(* Logix 5000 project; controller TFF vendor 1 type 14 code 107 rev 34.11; software revision 34.03; part 27 of 36 *)
(* tags used below, declared in another part *)
   BufferSteps0_Prev : STRING25;
   Config : Configuration;   // Index Array used in configuration routines
   Index : DINT;   // Index
   RecipeStepLog_DateTime_Empty : STRING25;   // Empty String
   RecipeStepLog_DateTime_Log : STRING25;   // Last Date Time received from HMI
   RecipeStepLog_DateTime_Prev : STRING25;
   RecipeStepLog_Timer : TIMER;   // RecipeStepLog Watchdog Timer
   AI101 : ALIAS FOR AnalogPoint[10];   // Filtrate Conductivity
   AI101_SIG : ALIAS FOR DigitalPoint[90];
   AI102 : ALIAS FOR AnalogPoint[11];   // Filtrate UV
   AI102_SIG : ALIAS FOR DigitalPoint[91];
   AI103 : ALIAS FOR AnalogPoint[12];   // Filtrate UV
   AI103_SIG : ALIAS FOR DigitalPoint[92];
   AI104 : ALIAS FOR AnalogPoint[9];   // Filtrate pH
   AI104_SIG : ALIAS FOR DigitalPoint[105];
   CCPSystem : CCPSystem;   // CCP System Data
   DigitalInput : BOOL[256];   // Digital Input Array these bits are copied from Input cards.
   DigitalPoint : DigitalPoint[150];   // Digital Point Array
   ES001 : ALIAS FOR DigitalPoint[3];   // Emergency Stop
   FI003 : ALIAS FOR AnalogPoint[17];
   FI003_SIG : ALIAS FOR DigitalPoint[106];
   FI101 : ALIAS FOR AnalogPoint[2];   // Filtrate Flow
   FI101_SIG : ALIAS FOR DigitalPoint[93];
   HTCCollectorError : BOOL;   // Hist. Data Collect. Error
   HTCHeartBeat : BOOL;   // Historical Data Collection heartbeat (Set to 1 by HMI Reset to 0 by PLC)
   MIX001 : ALIAS FOR AnalogPoint[14];   // Mixer Speed
   MIX001_SIG : ALIAS FOR DigitalPoint[104];
   Mixer : Mixer;   // Mixer config. structure
   OperatingTime : OperatingTime;
   Options : Options;   // Options List
   PcToPLCHeartBeat : BOOL;   // PC to PLC communication heartbeat Set to 1 by HMI Reset to 0 by plc
   PCV001 : ALIAS FOR AnalogPoint[3];   // Retentate Pressure Control Valve Position
   PCV001_SIG : ALIAS FOR DigitalPoint[102];
   PCV101 : ALIAS FOR AnalogPoint[4];   // Filtrate Pressure Control Valve Position
   PCV101_SIG : ALIAS FOR DigitalPoint[103];
   Phase0 : ALIAS FOR Phase[0];   // Phase 0
   PI001 : ALIAS FOR AnalogPoint[5];   // Feed Pressure
   PI001_SIG : ALIAS FOR DigitalPoint[97];
   PI002 : ALIAS FOR AnalogPoint[6];   // Retentate Pressure
   PI002_SIG : ALIAS FOR DigitalPoint[98];
   PI101 : ALIAS FOR AnalogPoint[7];   // Filtrate Pressure
   PI101_SIG : ALIAS FOR DigitalPoint[99];
   PI401 : ALIAS FOR AnalogPoint[8];   // Transfer Pump Pressure
   PI401_SIG : ALIAS FOR DigitalPoint[100];
   PSH001 : ALIAS FOR DigitalPoint[4];   // Feed Pump High Pressure
   PSH401 : ALIAS FOR DigitalPoint[5];   // Transfer Pump High Pressure
   PSL603 : ALIAS FOR DigitalPoint[10];   // Manifold Valves Air Defect
   Rack_Murr_Node0_Smart : IO_Station;   // Status of Node 0 Smart
   Rack_Murr_Node1_TF2S : IO_Station;   // Status of Node 1 TF2S
   Rack_Murr_Node1_TF3S : IO_Station;   // Status of Node 1 TF3S
   Rack_Murr_Node3_PUMP : IO_Station;   // Status of Node 3 Pump
   Rack_Murr_Node4_Instrum_TFF1 : IO_Station;   // Status of Node 4 Instrum TFF1
   Rack_Murr_Node4_Instrum_TFF2 : IO_Station;   // Status of Node 4 Instrum TFF2
   Rack_Murr_Node4_Instrum_TFF3 : IO_Station;   // Status of Node 4 Instrum TFF3
   Rack_Murr_Node4_Instrum_TFF4 : IO_Station;   // Status of Node 4 Instrum TFF4
   Rack_Murr_Node4_Instrum_TFF5 : IO_Station;   // Status of Node 4 Instrum TFF5
   Rack_Murr_Node5_Tank100 : IO_Station;   // Status of Node 5 Tank 100L
   Rack_Murr_Node5_Tank250 : IO_Station;   // Status of Node 5 Tank 250L
   Rack_Murr_Node5_Tank50 : IO_Station;   // Status of Node 5 Tank 50L
   Rack_Murr_Node6_IND331_WI001 : IO_Station;   // Status of Node 6 IND331 WI001
   Rack_Murr_Node7_IND131_WI101 : IO_Station;   // Status of Node 7 IND131 WI101
   RecipeStepLog_DateTime : STRING25;
   SIC001DF : ALIAS FOR DigitalPoint[8];   // Feed Pump Defect
   SIC002DF : ALIAS FOR DigitalPoint[9];   // Transfer Pump Defect
   SIC003DF : ALIAS FOR DigitalPoint[14];   // Mixer Defect
   SRL001 : ALIAS FOR DigitalPoint[15];   // Tank Skid Remote / Standalone
   Tank : TankManagement;   // Tank Management
   ThisSystem : SystemType;
   TI001 : ALIAS FOR AnalogPoint[13];   // Feed Bag Temperature
   TI001_SIG : ALIAS FOR DigitalPoint[101];
   WI001 : ALIAS FOR AnalogPoint[15];   // Feed Bag Weight
   WI001_SIG : ALIAS FOR DigitalPoint[94];
   WI101 : ALIAS FOR AnalogPoint[0];   // Filtrate Weight
   WI101_SIG : ALIAS FOR DigitalPoint[95];
   WI102 : ALIAS FOR AnalogPoint[1];   // Customer Filtrate Weight
   WI102_SIG : ALIAS FOR DigitalPoint[96];
   XC102_3DF : ALIAS FOR DigitalPoint[13];   // C8000 Defect
   XS001 : ALIAS FOR DigitalPoint[1];   // Door Closed
   XS002 : ALIAS FOR DigitalPoint[6];   // Clamshell Locking 1 Closed
   XS003 : ALIAS FOR DigitalPoint[7];   // Clamshell Locking 2 Closed
   XS006 : ALIAS FOR DigitalPoint[2];   // Door to Frame Locking Closed
   XS011 : ALIAS FOR DigitalPoint[11];   // Pump P001 Type
   XS012 : ALIAS FOR DigitalPoint[12];   // Pump P002 Type
   YA01 : ALIAS FOR DigitalPoint[50];   // PC to PLC communication failure
   YA02 : ALIAS FOR DigitalPoint[51];   // CCP Runtime communication failure
   YA03 : ALIAS FOR DigitalPoint[52];   // Historical Data collection failure
   YA06 : ALIAS FOR DigitalPoint[55];   // Node 0 communication failure - Smart
   YA07 : ALIAS FOR DigitalPoint[56];   // Node 0 internal defect - Smart
   YA08 : ALIAS FOR DigitalPoint[57];   // Node 1 communication failure - Clamshell
   YA09 : ALIAS FOR DigitalPoint[58];   // Node 1 internal defect - Clamshell
   YA13 : ALIAS FOR DigitalPoint[62];   // Tank Size Mismatch
   YA14 : ALIAS FOR DigitalPoint[63];   // SQL Server Write Failure
   YA15 : ALIAS FOR DigitalPoint[69];   // Node 3 Communication Failure - Pump
   YA16 : ALIAS FOR DigitalPoint[70];   // Node 3 Internal Defect - Pump
   YA17 : ALIAS FOR DigitalPoint[71];   // Node 4 Communication Failure - Instrum
   YA18 : ALIAS FOR DigitalPoint[72];   // Node 4 Internal Defect - Instrum
   YA19 : ALIAS FOR DigitalPoint[73];   // Node 5 Communication Failure - Tank
   YA20 : ALIAS FOR DigitalPoint[74];   // Node 5 Internal Defect - Tank
   YA21 : ALIAS FOR DigitalPoint[75];   // Node 6 IND331 Communication Failure
   YA22 : ALIAS FOR DigitalPoint[76];   // Node 7 IND131 Communication Failure
   YA41 : ALIAS FOR DigitalPoint[77];   // YA41 Operating Time Exceeded
   ZSDF : ALIAS FOR DigitalPoint[68];   // ZSDF Clamshell Locking Defect
(* Process, continued *)

ROUTINE InputDigitalPoint   (* ladder *)
// Digital Point Routine
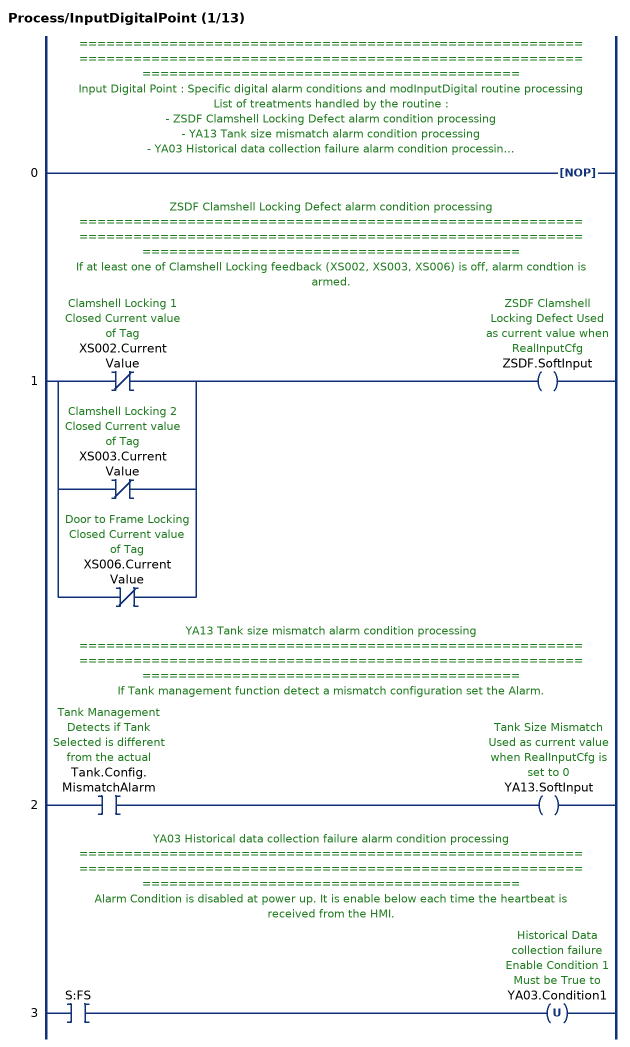
   // ==========================================================================================================================================================
   //                                                                                   Input Digital Point : Specific digital alarm conditions and modInputDigital routine processing
   //                                                     List of treatments handled by the routine :
   //                                                          - ZSDF Clamshell Locking Defect alarm condition processing
   //                                                          - YA13 Tank size mismatch alarm condition processing
   //                                                          - YA03 Historical data collection failure alarm condition processing
   //                                                          - YA01 PC to PLC com. failure alarm condition processing
   //                                                          - YA02 CCP Runtime com. failure alarm condition processing
   //                                                          - YA14 SQL Write failure alarm condition processing
   //                                                          - Node 0 communication failure and internal defect (YA06 and YA07)
   //                                                          - Node 1 communication failure and internal defect (YA08 and YA09)
   //                                                          - Node 3 communication failure and internal defect (YA15 and YA16)
   //                                                          - Node 4 communication failure and internal defect (YA17 and YA18)
   //                                                          - Node 5 communication failure and internal defect (YA19 and YA20)
   //                                                          - IND331 communication failure and internal defect (YA21)
   //                                                          - IND131 communication failure and internal defect (YA22)
   //                               - YA41 Operating Time Exceeded (YA41)
   //                                                          - Analog Signal Failure
   //                                                          - modInputDigital Loop
   //                                                     -----------------------------------------------------------------------------------------------------------------------------------------------------
   //                                                     History
   //                                            2019-AUG-13 - Actemium - B. Roch - Initial version for Candidate Release 3.00.00.00.a
   //                              2019-SEP-25 - Actemium - B. Roch - Modification for Candidate Release 3.00.00.00
   // - Add condition to comput SQL Write failure alarm (not in step 1)
   //                                 2020-SEP-14 - Merck - Q. Spindler - Modifications for Candidate Release 3.00.00.01.a
   //                                                   - Add Conditions to YA20, YA18, and YA09 so only connected nodes can trigger internal deffect
   //  - Change YA14 Alarm condition processing to add HMI Watchdog
   // - Add FI003_SIG
   // 2021-MAY-28 - DAVIDSON- Ch. ARBOGAST - Modifications for Candidate Release 3.01.00.00.a
   //  - Rung 6 unlatch YA03: add test not HTCColletorError (new tag - bool)
   //  - Add rung 30: write YA41.softInput - DigitalPoint[77] - Operating Time Exceeded
   // 2023-MAR-29 - DAVIDSON- Ch. ARBOGAST - Modifications for Candidate Release 3.02.00.00.a
   //  - Rung 2; replace DigitalPoint[41].SoftInput by YA13.SoftInput
   // ==========================================================================================================================================================
   0: NOP();
   // ZSDF Clamshell Locking Defect alarm condition processing
   // ==========================================================================================================================================================
   // If at least one of Clamshell Locking feedback (XS002, XS003, XS006) is off, alarm condtion is armed.
   1: [XIO(XS002.CurrentValue) ,XIO(XS003.CurrentValue) ,XIO(XS006.CurrentValue) ]OTE(ZSDF.SoftInput);
   // YA13 Tank size mismatch alarm condition processing
   // ==========================================================================================================================================================
   // If Tank management function detect a mismatch configuration set the Alarm.
   2: XIC(Tank.Config.MismatchAlarm)OTE(YA13.SoftInput);
   // YA03 Historical data collection failure alarm condition processing
   // ==========================================================================================================================================================
   // Alarm Condition is disabled at power up. It is enable below each time the heartbeat is received from the HMI.
   3: XIC(S:FS)OTU(YA03.Condition1);
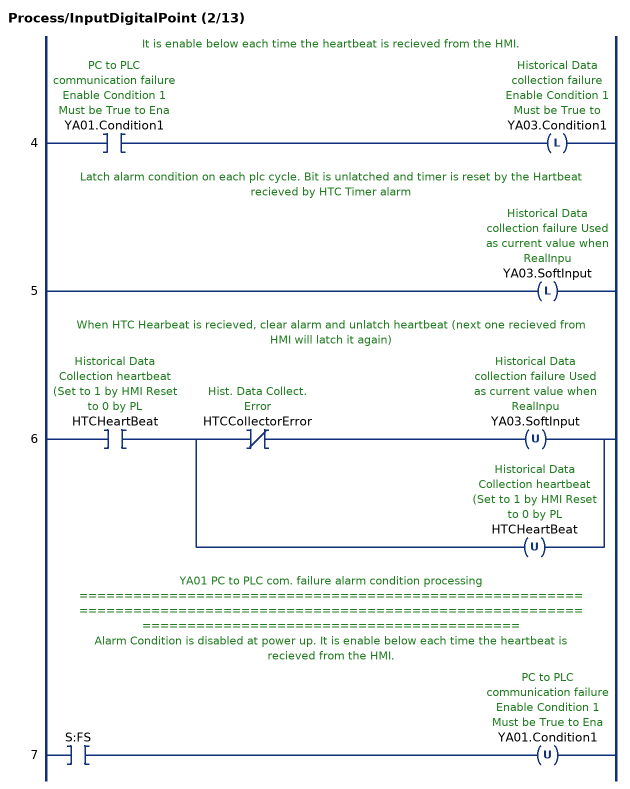
   // It is enable below each time the heartbeat is recieved from the HMI.
   4: XIC(YA01.Condition1)OTL(YA03.Condition1);
   // Latch alarm condition on each plc cycle. Bit is unlatched and timer is reset by the Hartbeat recieved by HTC Timer alarm
   5: OTL(YA03.SoftInput);
   // When HTC Hearbeat is recieved, clear alarm and unlatch heartbeat (next one recieved from HMI will latch it again)
   6: XIC(HTCHeartBeat)[XIO(HTCCollectorError) OTU(YA03.SoftInput) ,OTU(HTCHeartBeat) ];
   // YA01 PC to PLC com. failure alarm condition processing
   // ==========================================================================================================================================================
   // Alarm Condition is disabled at power up. It is enable below each time the heartbeat is recieved from the HMI.
   7: XIC(S:FS)OTU(YA01.Condition1);
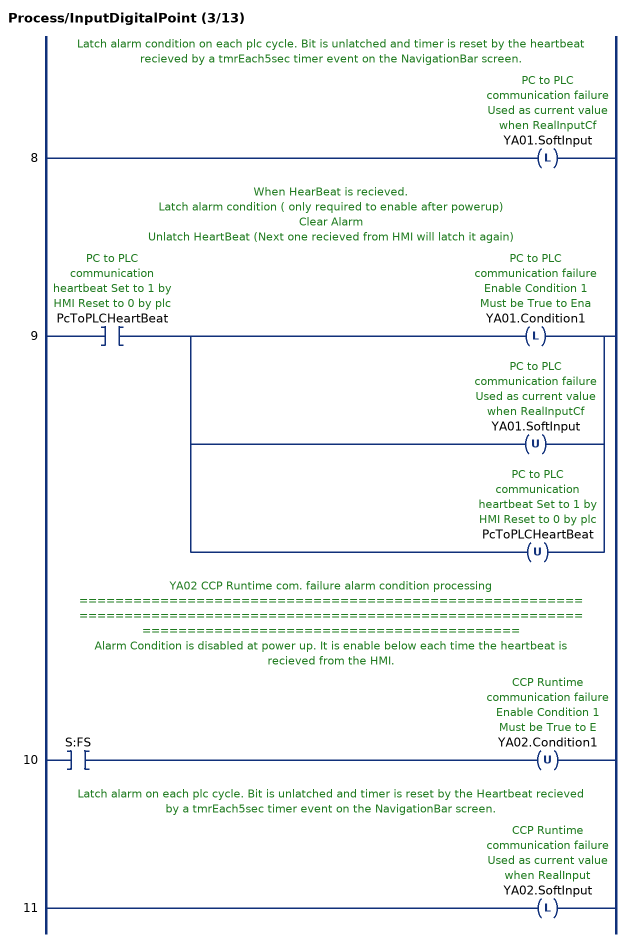
   // Latch alarm condition on each plc cycle. Bit is unlatched and timer is reset by the heartbeat recieved by a tmrEach5sec timer event on the NavigationBar screen.
   8: OTL(YA01.SoftInput);
   // When HearBeat is recieved.
   //         Latch alarm condition ( only required to enable after powerup)
   //         Clear Alarm
   //        Unlatch HeartBeat (Next one recieved from HMI will latch it again)
   9: XIC(PcToPLCHeartBeat)[OTL(YA01.Condition1) ,OTU(YA01.SoftInput) ,OTU(PcToPLCHeartBeat) ];
   // YA02 CCP Runtime com. failure alarm condition processing
   // ==========================================================================================================================================================
   // Alarm Condition is disabled at power up. It is enable below each time the heartbeat is recieved from the HMI.
   10: XIC(S:FS)OTU(YA02.Condition1);
   // Latch alarm on each plc cycle. Bit is unlatched and timer is reset by the Heartbeat recieved by a tmrEach5sec timer event on the NavigationBar screen.
   11: OTL(YA02.SoftInput);
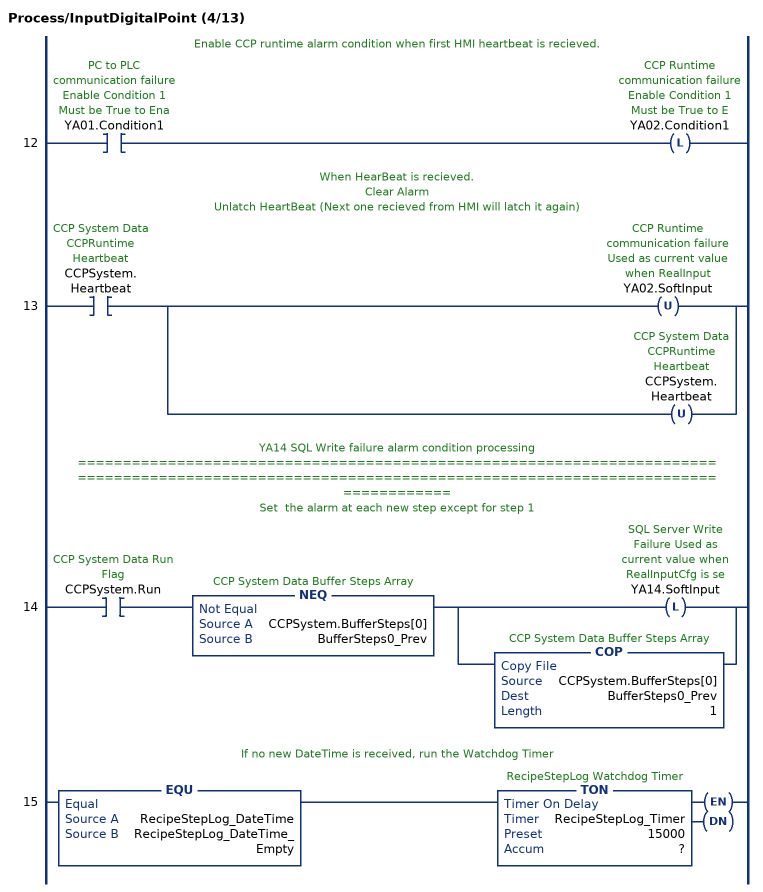
   // Enable CCP runtime alarm condition when first HMI heartbeat is recieved.
   12: XIC(YA01.Condition1)OTL(YA02.Condition1);
   // When HearBeat is recieved.
   //         Clear Alarm
   //        Unlatch HeartBeat (Next one recieved from HMI will latch it again)
   13: XIC(CCPSystem.Heartbeat)[OTU(YA02.SoftInput) ,OTU(CCPSystem.Heartbeat) ];
   // YA14 SQL Write failure alarm condition processing
   // ==========================================================================================================================================================
   // Set  the alarm at each new step except for step 1
   14: XIC(CCPSystem.Run)NEQ(CCPSystem.BufferSteps[0],BufferSteps0_Prev)[OTL(YA14.SoftInput) ,COP(CCPSystem.BufferSteps[0],BufferSteps0_Prev,1) ];
   // If no new DateTime is received, run the Watchdog Timer
   15: EQU(RecipeStepLog_DateTime,RecipeStepLog_DateTime_Empty)TON(RecipeStepLog_Timer,?,?);
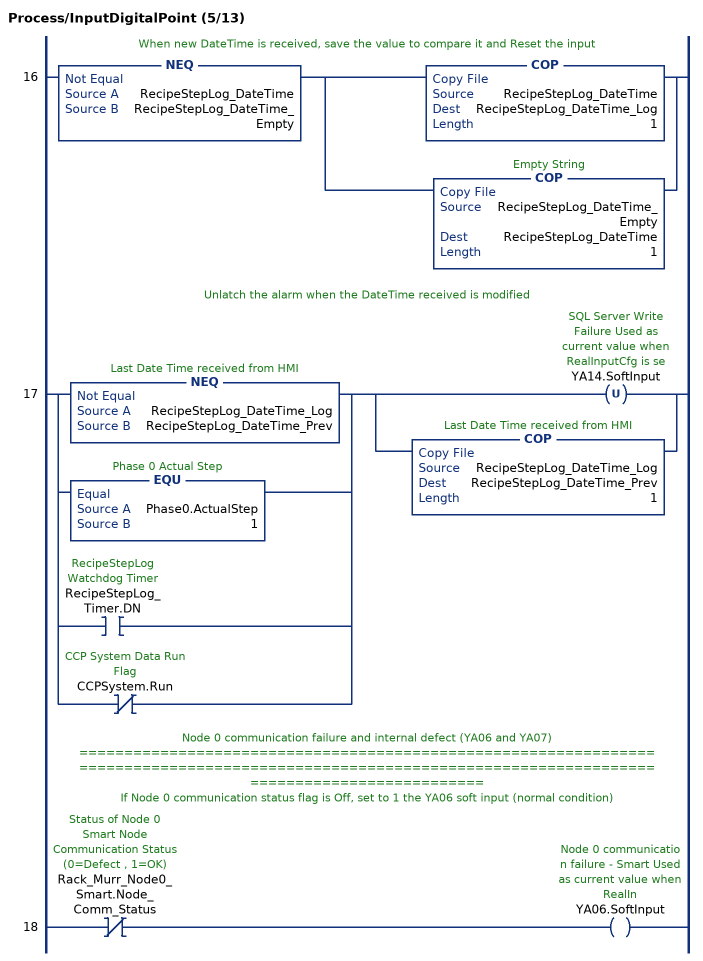
   // When new DateTime is received, save the value to compare it and Reset the input
   16: NEQ(RecipeStepLog_DateTime,RecipeStepLog_DateTime_Empty)[COP(RecipeStepLog_DateTime,RecipeStepLog_DateTime_Log,1) ,COP(RecipeStepLog_DateTime_Empty,RecipeStepLog_DateTime,1) ];
   // Unlatch the alarm when the DateTime received is modified
   17: [NEQ(RecipeStepLog_DateTime_Log,RecipeStepLog_DateTime_Prev) ,EQU(Phase0.ActualStep,1) ,XIC(RecipeStepLog_Timer.DN) ,XIO(CCPSystem.Run) ][OTU(YA14.SoftInput) ,COP(RecipeStepLog_DateTime_Log,RecipeStepLog_DateTime_Prev,1) ];
   // Node 0 communication failure and internal defect (YA06 and YA07)
   // ==========================================================================================================================================================
   // If Node 0 communication status flag is Off, set to 1 the YA06 soft input (normal condition)
   18: XIO(Rack_Murr_Node0_Smart.Node_Comm_Status)OTE(YA06.SoftInput);
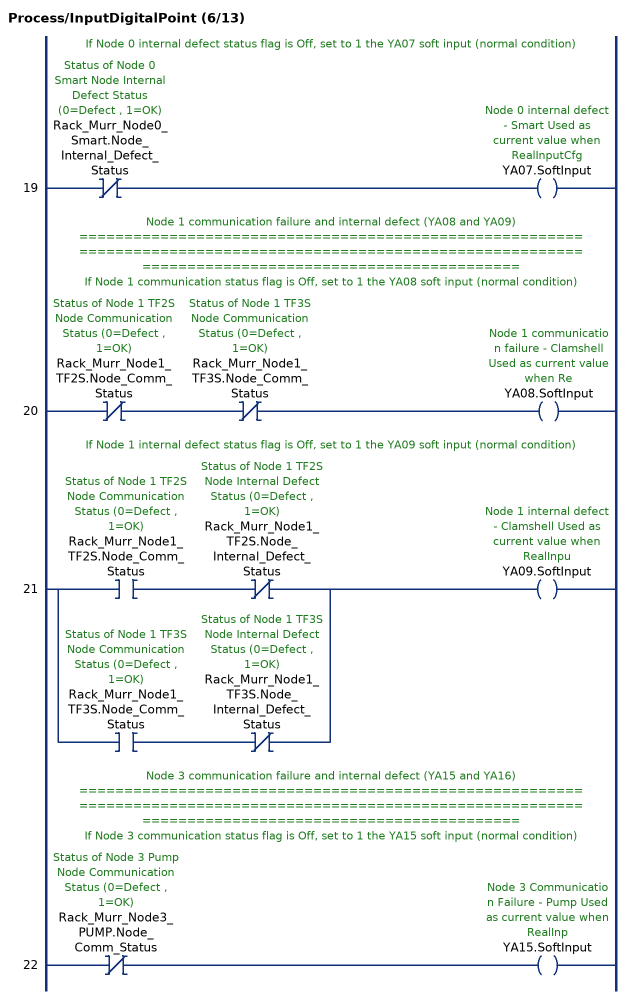
   // If Node 0 internal defect status flag is Off, set to 1 the YA07 soft input (normal condition)
   19: XIO(Rack_Murr_Node0_Smart.Node_Internal_Defect_Status)OTE(YA07.SoftInput);
   // Node 1 communication failure and internal defect (YA08 and YA09)
   // ==========================================================================================================================================================
   // If Node 1 communication status flag is Off, set to 1 the YA08 soft input (normal condition)
   20: XIO(Rack_Murr_Node1_TF2S.Node_Comm_Status)XIO(Rack_Murr_Node1_TF3S.Node_Comm_Status)OTE(YA08.SoftInput);
   // If Node 1 internal defect status flag is Off, set to 1 the YA09 soft input (normal condition)
   21: [XIC(Rack_Murr_Node1_TF2S.Node_Comm_Status) XIO(Rack_Murr_Node1_TF2S.Node_Internal_Defect_Status) ,XIC(Rack_Murr_Node1_TF3S.Node_Comm_Status) XIO(Rack_Murr_Node1_TF3S.Node_Internal_Defect_Status) ]OTE(YA09.SoftInput);
   // Node 3 communication failure and internal defect (YA15 and YA16)
   // ==========================================================================================================================================================
   // If Node 3 communication status flag is Off, set to 1 the YA15 soft input (normal condition)
   22: XIO(Rack_Murr_Node3_PUMP.Node_Comm_Status)OTE(YA15.SoftInput);
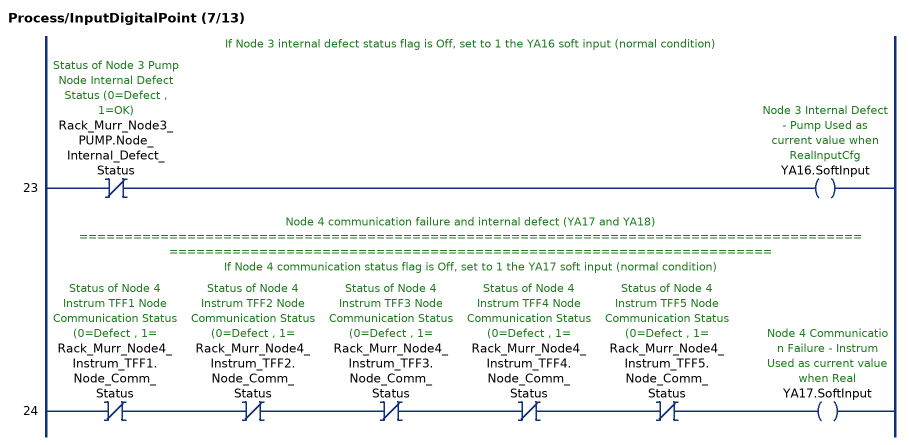
   // If Node 3 internal defect status flag is Off, set to 1 the YA16 soft input (normal condition)
   23: XIO(Rack_Murr_Node3_PUMP.Node_Internal_Defect_Status)OTE(YA16.SoftInput);
   // Node 4 communication failure and internal defect (YA17 and YA18)
   // ==========================================================================================================================================================
   // If Node 4 communication status flag is Off, set to 1 the YA17 soft input (normal condition)
   24: XIO(Rack_Murr_Node4_Instrum_TFF1.Node_Comm_Status)XIO(Rack_Murr_Node4_Instrum_TFF2.Node_Comm_Status)XIO(Rack_Murr_Node4_Instrum_TFF3.Node_Comm_Status)XIO(Rack_Murr_Node4_Instrum_TFF4.Node_Comm_Status)XIO(Rack_Murr_Node4_Instrum_TFF5.Node_Comm_Status)OTE(YA17.SoftInput);
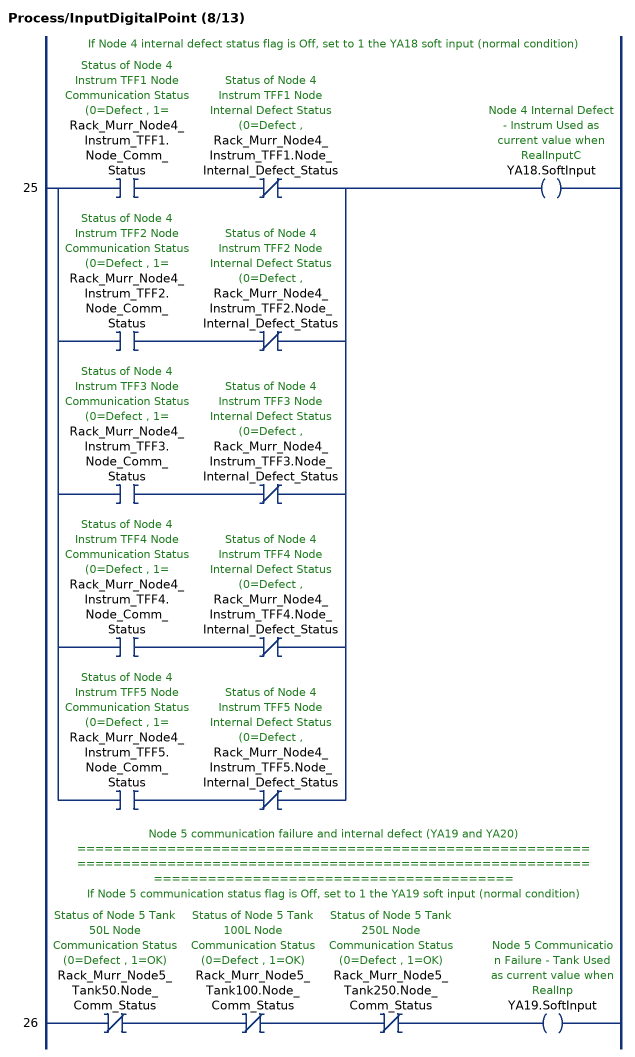
   // If Node 4 internal defect status flag is Off, set to 1 the YA18 soft input (normal condition)
   25: [XIC(Rack_Murr_Node4_Instrum_TFF1.Node_Comm_Status) XIO(Rack_Murr_Node4_Instrum_TFF1.Node_Internal_Defect_Status) ,XIC(Rack_Murr_Node4_Instrum_TFF2.Node_Comm_Status) XIO(Rack_Murr_Node4_Instrum_TFF2.Node_Internal_Defect_Status) ,XIC(Rack_Murr_Node4_Instrum_TFF3.Node_Comm_Status) XIO(Rack_Murr_Node4_Instrum_TFF3.Node_Internal_Defect_Status) ,XIC(Rack_Murr_Node4_Instrum_TFF4.Node_Comm_Status) XIO(Rack_Murr_Node4_Instrum_TFF4.Node_Internal_Defect_Status) ,XIC(Rack_Murr_Node4_Instrum_TFF5.Node_Comm_Status) XIO(Rack_Murr_Node4_Instrum_TFF5.Node_Internal_Defect_Status) ]OTE(YA18.SoftInput);
   // Node 5 communication failure and internal defect (YA19 and YA20)
   // ==========================================================================================================================================================
   // If Node 5 communication status flag is Off, set to 1 the YA19 soft input (normal condition)
   26: XIO(Rack_Murr_Node5_Tank50.Node_Comm_Status)XIO(Rack_Murr_Node5_Tank100.Node_Comm_Status)XIO(Rack_Murr_Node5_Tank250.Node_Comm_Status)OTE(YA19.SoftInput);
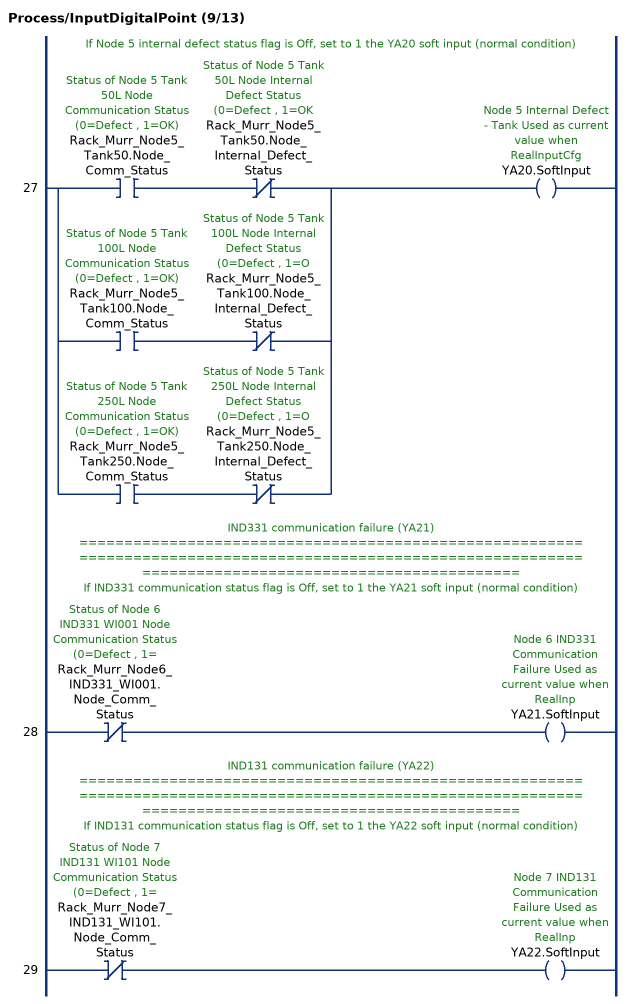
   // If Node 5 internal defect status flag is Off, set to 1 the YA20 soft input (normal condition)
   27: [XIC(Rack_Murr_Node5_Tank50.Node_Comm_Status) XIO(Rack_Murr_Node5_Tank50.Node_Internal_Defect_Status) ,XIC(Rack_Murr_Node5_Tank100.Node_Comm_Status) XIO(Rack_Murr_Node5_Tank100.Node_Internal_Defect_Status) ,XIC(Rack_Murr_Node5_Tank250.Node_Comm_Status) XIO(Rack_Murr_Node5_Tank250.Node_Internal_Defect_Status) ]OTE(YA20.SoftInput);
   // IND331 communication failure (YA21)
   // ==========================================================================================================================================================
   // If IND331 communication status flag is Off, set to 1 the YA21 soft input (normal condition)
   28: XIO(Rack_Murr_Node6_IND331_WI001.Node_Comm_Status)OTE(YA21.SoftInput);
   // IND131 communication failure (YA22)
   // ==========================================================================================================================================================
   // If IND131 communication status flag is Off, set to 1 the YA22 soft input (normal condition)
   29: XIO(Rack_Murr_Node7_IND131_WI101.Node_Comm_Status)OTE(YA22.SoftInput);
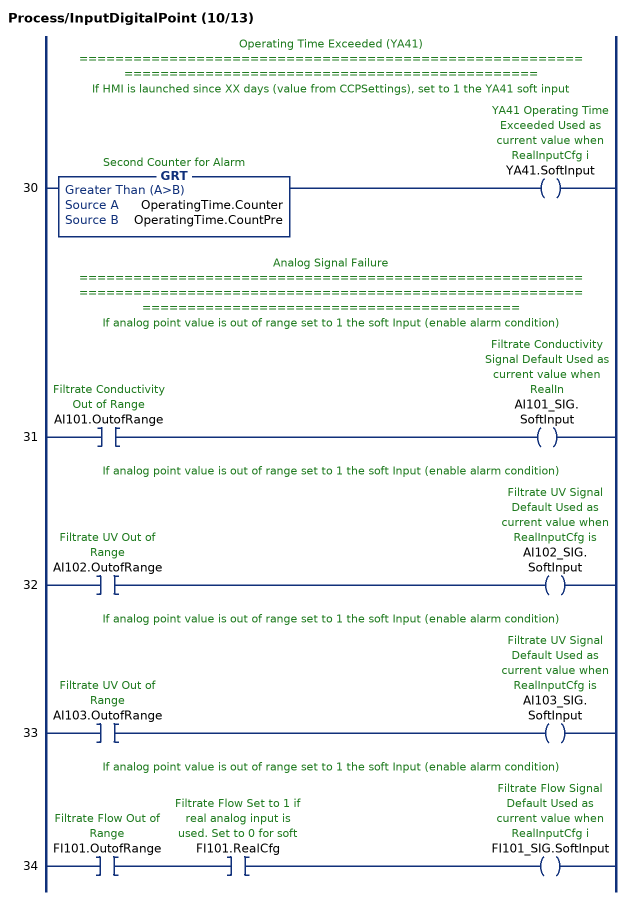
   // Operating Time Exceeded (YA41)
   // ======================================================================================================
   // If HMI is launched since XX days (value from CCPSettings), set to 1 the YA41 soft input
   30: GRT(OperatingTime.Counter,OperatingTime.CountPre)OTE(YA41.SoftInput);
   // Analog Signal Failure
   // ==========================================================================================================================================================
   // If analog point value is out of range set to 1 the soft Input (enable alarm condition)
   31: XIC(AI101.OutofRange)OTE(AI101_SIG.SoftInput);
   // If analog point value is out of range set to 1 the soft Input (enable alarm condition)
   32: XIC(AI102.OutofRange)OTE(AI102_SIG.SoftInput);
   // If analog point value is out of range set to 1 the soft Input (enable alarm condition)
   33: XIC(AI103.OutofRange)OTE(AI103_SIG.SoftInput);
   // If analog point value is out of range set to 1 the soft Input (enable alarm condition)
   34: XIC(FI101.OutofRange)XIC(FI101.RealCfg)OTE(FI101_SIG.SoftInput);
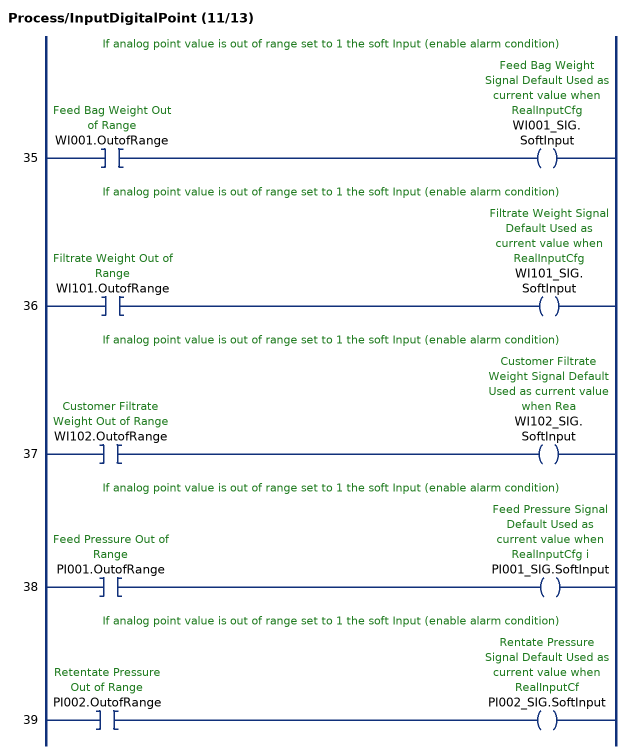
   // If analog point value is out of range set to 1 the soft Input (enable alarm condition)
   35: XIC(WI001.OutofRange)OTE(WI001_SIG.SoftInput);
   // If analog point value is out of range set to 1 the soft Input (enable alarm condition)
   36: XIC(WI101.OutofRange)OTE(WI101_SIG.SoftInput);
   // If analog point value is out of range set to 1 the soft Input (enable alarm condition)
   37: XIC(WI102.OutofRange)OTE(WI102_SIG.SoftInput);
   // If analog point value is out of range set to 1 the soft Input (enable alarm condition)
   38: XIC(PI001.OutofRange)OTE(PI001_SIG.SoftInput);
   // If analog point value is out of range set to 1 the soft Input (enable alarm condition)
   39: XIC(PI002.OutofRange)OTE(PI002_SIG.SoftInput);
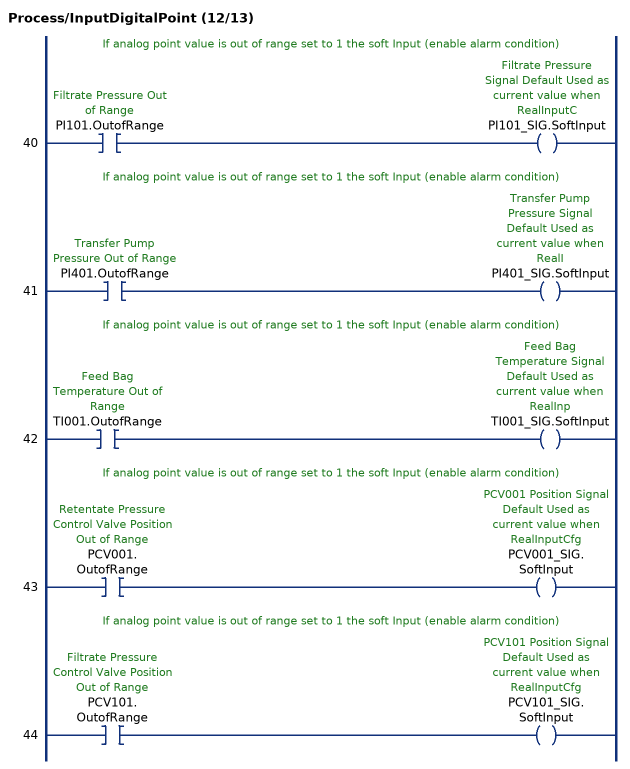
   // If analog point value is out of range set to 1 the soft Input (enable alarm condition)
   40: XIC(PI101.OutofRange)OTE(PI101_SIG.SoftInput);
   // If analog point value is out of range set to 1 the soft Input (enable alarm condition)
   41: XIC(PI401.OutofRange)OTE(PI401_SIG.SoftInput);
   // If analog point value is out of range set to 1 the soft Input (enable alarm condition)
   42: XIC(TI001.OutofRange)OTE(TI001_SIG.SoftInput);
   // If analog point value is out of range set to 1 the soft Input (enable alarm condition)
   43: XIC(PCV001.OutofRange)OTE(PCV001_SIG.SoftInput);
   // If analog point value is out of range set to 1 the soft Input (enable alarm condition)
   44: XIC(PCV101.OutofRange)OTE(PCV101_SIG.SoftInput);
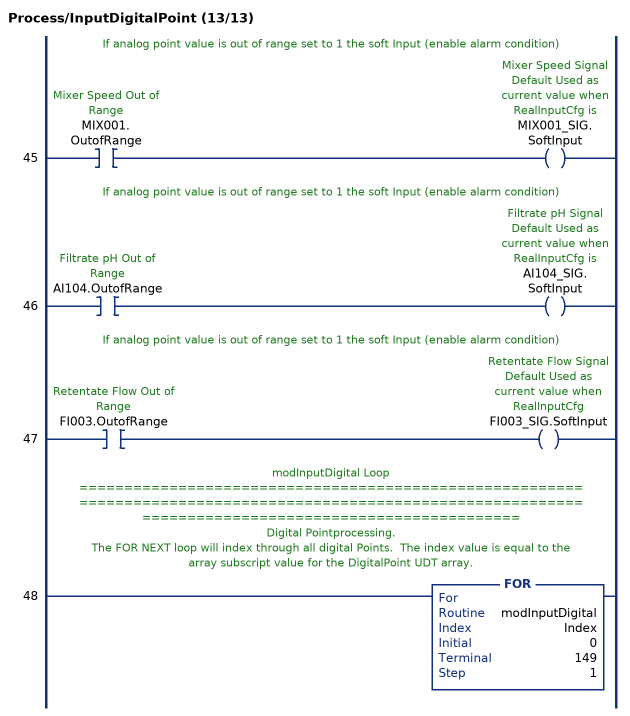
   // If analog point value is out of range set to 1 the soft Input (enable alarm condition)
   45: XIC(MIX001.OutofRange)OTE(MIX001_SIG.SoftInput);
   // If analog point value is out of range set to 1 the soft Input (enable alarm condition)
   46: XIC(AI104.OutofRange)OTE(AI104_SIG.SoftInput);
   // If analog point value is out of range set to 1 the soft Input (enable alarm condition)
   47: XIC(FI003.OutofRange)OTE(FI003_SIG.SoftInput);
   // modInputDigital Loop
   // ==========================================================================================================================================================
   // Digital Pointprocessing.
   // The FOR NEXT loop will index through all digital Points.  The index value is equal to the array subscript value for the DigitalPoint UDT array.
   48: FOR(modInputDigital,Index,0,149,1);
END_ROUTINE

ROUTINE InputDigitalRaw   (* ladder *)
// Digital Input Routine
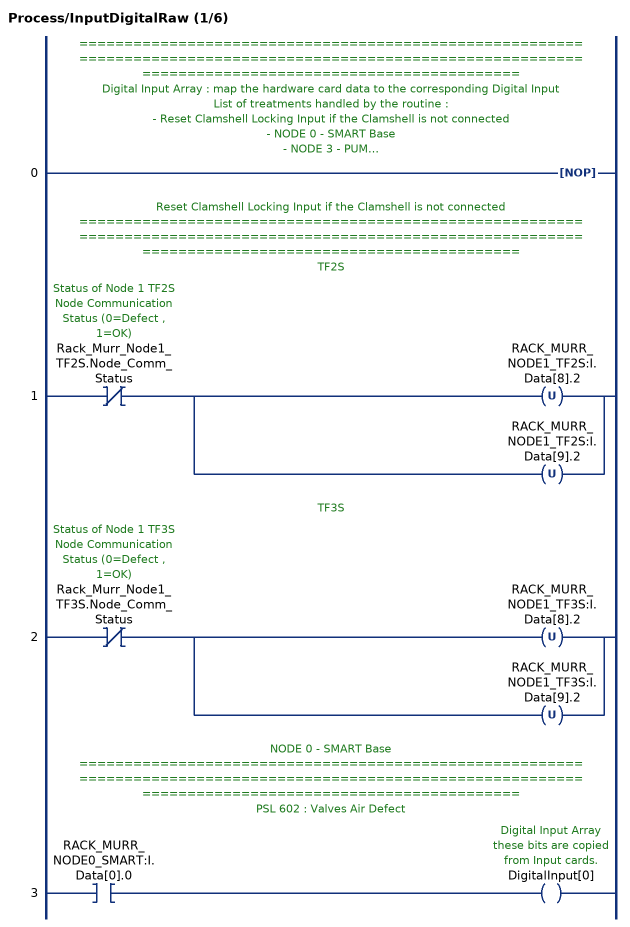
   // ==========================================================================================================================================================
   //                                                                                             Digital Input Array : map the hardware card data to the corresponding Digital Input
   //                                                     List of treatments handled by the routine :
   //                                                    - Reset Clamshell Locking Input if the Clamshell is not connected
   //                                                    - NODE 0 - SMART Base
   //                                                    - NODE 3 - PUMP
   //                                                    - NODE 4 - INSTRUM
   //                                                    - NODE 5 - TANK
   //                                                    - NODE 1 - TF2S
   //                                                    - NODE 1 - TF3S
   //                                                     -----------------------------------------------------------------------------------------------------------------------------------------------------
   //                                                     History
   //                                                          2019-AUG-13 - Actemium - B. Roch - Initial version for Candidate Release 3.00.00.00.a
   // ==========================================================================================================================================================
   0: NOP();
   // Reset Clamshell Locking Input if the Clamshell is not connected
   // ==========================================================================================================================================================
   // TF2S
   1: XIO(Rack_Murr_Node1_TF2S.Node_Comm_Status)[OTU(RACK_MURR_NODE1_TF2S:I.Data[8].2) ,OTU(RACK_MURR_NODE1_TF2S:I.Data[9].2) ];
   // TF3S
   2: XIO(Rack_Murr_Node1_TF3S.Node_Comm_Status)[OTU(RACK_MURR_NODE1_TF3S:I.Data[8].2) ,OTU(RACK_MURR_NODE1_TF3S:I.Data[9].2) ];
   // NODE 0 - SMART Base
   // ==========================================================================================================================================================
   // PSL 602 : Valves Air Defect
   3: XIC(RACK_MURR_NODE0_SMART:I.Data[0].0)OTE(DigitalInput[0]);
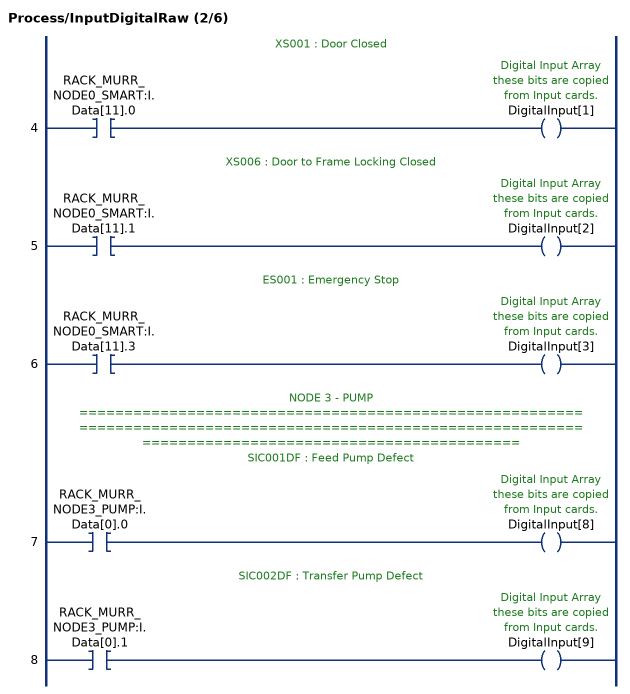
   // XS001 : Door Closed
   4: XIC(RACK_MURR_NODE0_SMART:I.Data[11].0)OTE(DigitalInput[1]);
   // XS006 : Door to Frame Locking Closed
   5: XIC(RACK_MURR_NODE0_SMART:I.Data[11].1)OTE(DigitalInput[2]);
   // ES001 : Emergency Stop
   6: XIC(RACK_MURR_NODE0_SMART:I.Data[11].3)OTE(DigitalInput[3]);
   // NODE 3 - PUMP
   // ==========================================================================================================================================================
   // SIC001DF : Feed Pump Defect
   7: XIC(RACK_MURR_NODE3_PUMP:I.Data[0].0)OTE(DigitalInput[8]);
   // SIC002DF : Transfer Pump Defect
   8: XIC(RACK_MURR_NODE3_PUMP:I.Data[0].1)OTE(DigitalInput[9]);
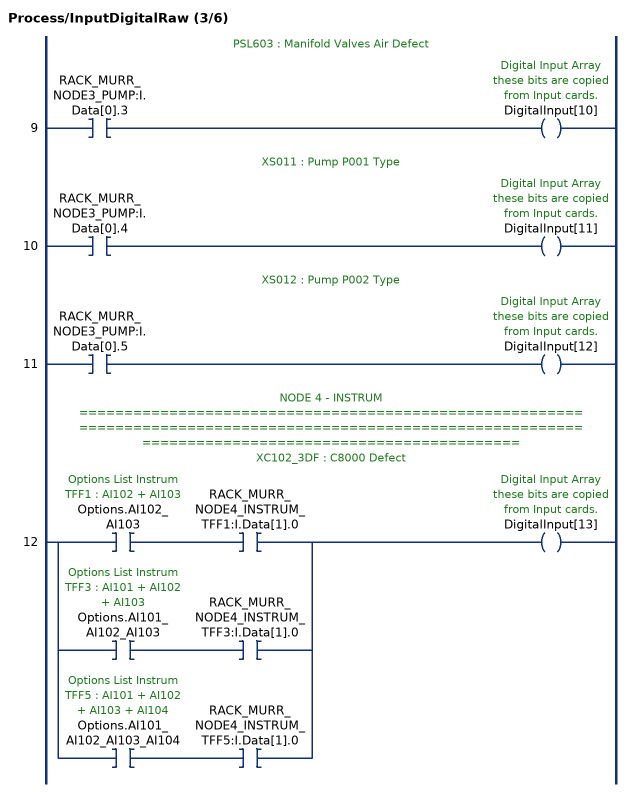
   // PSL603 : Manifold Valves Air Defect
   9: XIC(RACK_MURR_NODE3_PUMP:I.Data[0].3)OTE(DigitalInput[10]);
   // XS011 : Pump P001 Type
   10: XIC(RACK_MURR_NODE3_PUMP:I.Data[0].4)OTE(DigitalInput[11]);
   // XS012 : Pump P002 Type
   11: XIC(RACK_MURR_NODE3_PUMP:I.Data[0].5)OTE(DigitalInput[12]);
   // NODE 4 - INSTRUM
   // ==========================================================================================================================================================
   // XC102_3DF : C8000 Defect
   12: [XIC(Options.AI102_AI103) XIC(RACK_MURR_NODE4_INSTRUM_TFF1:I.Data[1].0) ,XIC(Options.AI101_AI102_AI103) XIC(RACK_MURR_NODE4_INSTRUM_TFF3:I.Data[1].0) ,XIC(Options.AI101_AI102_AI103_AI104) XIC(RACK_MURR_NODE4_INSTRUM_TFF5:I.Data[1].0) ]OTE(DigitalInput[13]);
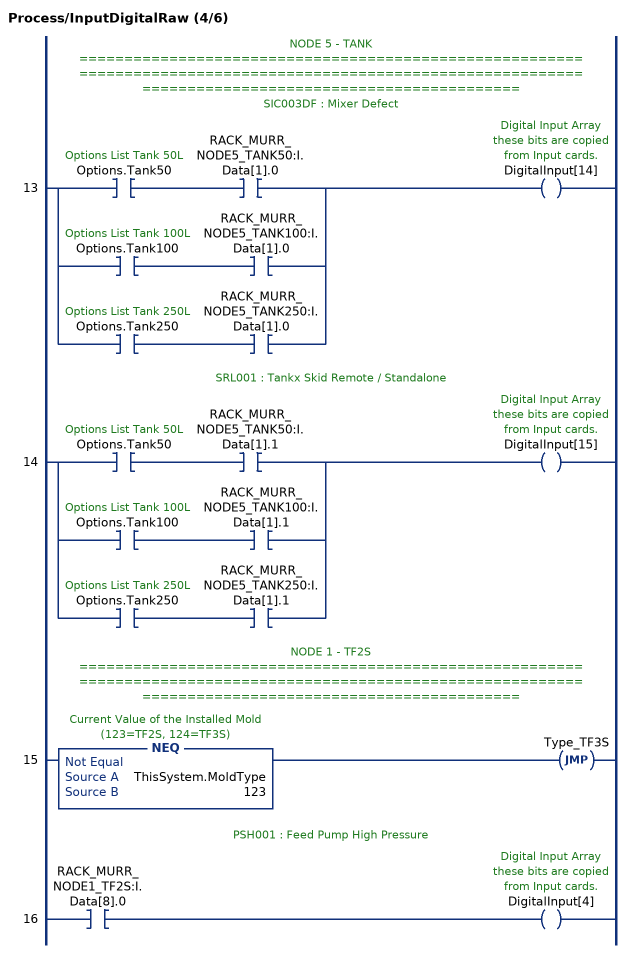
   // NODE 5 - TANK
   // ==========================================================================================================================================================
   // SIC003DF : Mixer Defect
   13: [XIC(Options.Tank50) XIC(RACK_MURR_NODE5_TANK50:I.Data[1].0) ,XIC(Options.Tank100) XIC(RACK_MURR_NODE5_TANK100:I.Data[1].0) ,XIC(Options.Tank250) XIC(RACK_MURR_NODE5_TANK250:I.Data[1].0) ]OTE(DigitalInput[14]);
   // SRL001 : Tankx Skid Remote / Standalone
   14: [XIC(Options.Tank50) XIC(RACK_MURR_NODE5_TANK50:I.Data[1].1) ,XIC(Options.Tank100) XIC(RACK_MURR_NODE5_TANK100:I.Data[1].1) ,XIC(Options.Tank250) XIC(RACK_MURR_NODE5_TANK250:I.Data[1].1) ]OTE(DigitalInput[15]);
   // NODE 1 - TF2S
   // ==========================================================================================================================================================
   15: NEQ(ThisSystem.MoldType,123)JMP(Type_TF3S);
   // PSH001 : Feed Pump High Pressure
   16: XIC(RACK_MURR_NODE1_TF2S:I.Data[8].0)OTE(DigitalInput[4]);
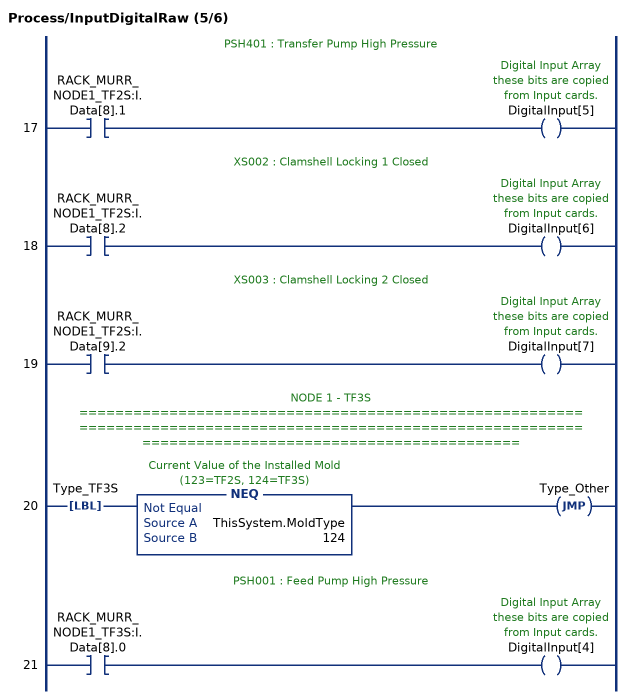
   // PSH401 : Transfer Pump High Pressure
   17: XIC(RACK_MURR_NODE1_TF2S:I.Data[8].1)OTE(DigitalInput[5]);
   // XS002 : Clamshell Locking 1 Closed
   18: XIC(RACK_MURR_NODE1_TF2S:I.Data[8].2)OTE(DigitalInput[6]);
   // XS003 : Clamshell Locking 2 Closed
   19: XIC(RACK_MURR_NODE1_TF2S:I.Data[9].2)OTE(DigitalInput[7]);
   // NODE 1 - TF3S
   // ==========================================================================================================================================================
   20: LBL(Type_TF3S)NEQ(ThisSystem.MoldType,124)JMP(Type_Other);
   // PSH001 : Feed Pump High Pressure
   21: XIC(RACK_MURR_NODE1_TF3S:I.Data[8].0)OTE(DigitalInput[4]);
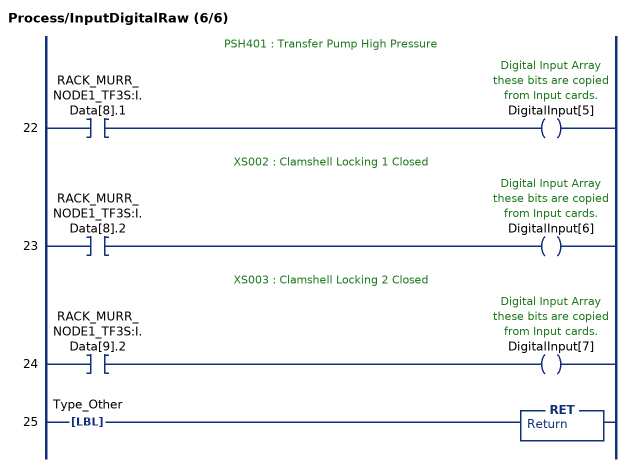
   // PSH401 : Transfer Pump High Pressure
   22: XIC(RACK_MURR_NODE1_TF3S:I.Data[8].1)OTE(DigitalInput[5]);
   // XS002 : Clamshell Locking 1 Closed
   23: XIC(RACK_MURR_NODE1_TF3S:I.Data[8].2)OTE(DigitalInput[6]);
   // XS003 : Clamshell Locking 2 Closed
   24: XIC(RACK_MURR_NODE1_TF3S:I.Data[9].2)OTE(DigitalInput[7]);
   25: LBL(Type_Other)RET();
END_ROUTINE
